Fanuc KAREL source: KT00805.KL

PROGRAM KT00805
%NOLOCKGROUP
VAR
  B1: BOOLEAN
  B2: BOOLEAN
  OUT: REAL
BEGIN
  B1 = TRUE
  B2 = FALSE
  B1 = TRUE
  B2 = FALSE
  OUT = EXP(B1)
END KT00805
